// TIA Portal V21 export
// export: Created 2026-11-11T00:47:22.7088143Z, ExportSetting WithDefaults, DisplayName Totally Integrated Automation Portal, DisplayVersion V21 Update 3, DisplayName STEP 7 Professional, DisplayVersion V21 Update 3, DisplayName STEP 7 Safety, DisplayVersion V21, DisplayName Tech WebApplication, DisplayVersion V21, DisplayName WinCC Basic/Comfort/Advanced, DisplayVersion V21 Update 3, DisplayName WinCC Unified, DisplayVersion V21 Update 3
FUNCTION_BLOCK "FB_Fbd_ex071"   // FB362, FBD
{ S7_Optimized_Access := 'TRUE' }
VERSION : 0.1
// stored: AutoNumber true, IsIECCheckEnabled false, IsRetainMemResEnabled false, MemoryReserve 100, SetENOAutomatically false, UDAEnableTagReadback false
   VAR_INPUT
      v_com_rst : Bool;
      v_start : Bool;
      v_end : Bool;
   END_VAR
   VAR_OUTPUT
      v_status : DWord;
   END_VAR
   VAR_IN_OUT
      v_penergy : PE_PLUS;
   END_VAR
   VAR
      inst { S7_SetPoint := 'True'} : PE_WOL;
   END_VAR
BEGIN

REGION Network 1: Description PE_WOL
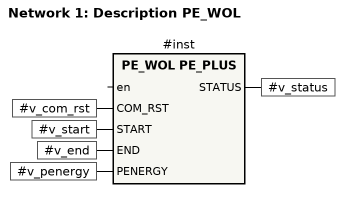
   #inst(COM_RST := #v_com_rst, START := #v_start, END := #v_end, PENERGY := #v_penergy, STATUS => #v_status);   // PE_WOL
END_REGION
END_FUNCTION_BLOCK
